(* PLC project Vn_fb_ctud, Beckhoff Automation GmbH TwinCAT PLC Control 3.5.13.21 *)
(* stored: creationDateTime 1970-01-01T00:00:00 *)

PROGRAM Vn_fb_ctud

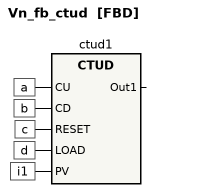
(* FBD diagram, written out as Structured Text *)
ctud1(CU := a, CD := b, RESET := c, LOAD := d, PV := i1);
END_PROGRAM
